// TIA Portal V21 export
// export: Created 2026-11-10T07:35:28.867292Z, ExportSetting WithDefaults, DisplayName Totally Integrated Automation Portal, DisplayVersion V21 Update 3, DisplayName STEP 7 Professional, DisplayVersion V21 Update 3, DisplayName STEP 7 Safety, DisplayVersion V21, DisplayName Tech WebApplication, DisplayVersion V21, DisplayName WinCC Basic/Comfort/Advanced, DisplayVersion V21 Update 3, DisplayName WinCC Unified, DisplayVersion V21 Update 3
FUNCTION_BLOCK "FB_Lad_sc006"   // FB88, LAD
{ S7_Optimized_Access := 'TRUE' }
VERSION : 0.1
// stored: AutoNumber true, IsIECCheckEnabled false, IsRetainMemResEnabled false, MemoryReserve 100, SetENOAutomatically false, UDAEnableTagReadback false
   VAR_INPUT
      v_en_r : Bool;
      v_id : CONN_PRG;
      v_r_id : CONN_R_ID;
   END_VAR
   VAR_OUTPUT
      v_ndr : Bool;
      v_error : Bool;
      v_status : Word;
   END_VAR
   VAR_IN_OUT
      v_rd_1 : Array[0..99] of Byte;
      v_len : Word;
   END_VAR
   VAR
      inst { S7_SetPoint := 'True'} : BRCV;
   END_VAR
BEGIN

REGION Network 1: BRCV - Receive data in segments
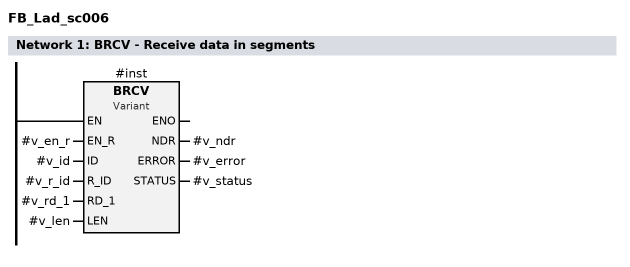
   RUNG wire#powerrail
      { S7_Templates := "[ptr_type := Variant, id_type := CONN_PRG, r_id_type := CONN_R_ID]" } #inst.BRCV(EN_R := #v_en_r, ID := #v_id, R_ID := #v_r_id, RD_1 := #v_rd_1, LEN := #v_len, NDR => #v_ndr, ERROR => #v_error, STATUS => #v_status)
   END_RUNG
   // the same network as SCL:
   #inst(EN_R := #v_en_r,   // BRCV
         ID := #v_id,
         R_ID := #v_r_id,
         RD_1 := #v_rd_1,
         LEN := #v_len,
         NDR => #v_ndr,
         ERROR => #v_error,
         STATUS => #v_status);
END_REGION
END_FUNCTION_BLOCK
